// TIA Portal V19 export
// export: Created 2026-10-15T09:44:25.0424598Z, ExportSetting WithDefaults, DisplayName Totally Integrated Automation Portal, DisplayVersion V19, DisplayName TIA Portal Openness, DisplayVersion V19, DisplayName TIA Portal Version Control Interface, DisplayVersion V19, DisplayName STEP 7 Professional, DisplayVersion V19, DisplayName STEP 7 Safety, DisplayVersion V19, DisplayName WinCC Basic/Comfort/Advanced, DisplayVersion V19, DisplayName WinCC Unified, DisplayVersion V19
FUNCTION "ROLL_PB52" : Void   // FC35, SCL
{ S7_Optimized_Access := 'TRUE' }
VERSION : 0.1
// stored: AutoNumber true, IsIECCheckEnabled false, SetENOAutomatically false, UDAEnableTagReadback false
   VAR_TEMP
      r : Bool;
      a1 : Word;
      a2 : Word;
      activeDataBlock : Int;
      comparisonResults : Array[0..0] of Bool;
   END_VAR
BEGIN

   #r := FALSE;
   #a1 := W#16#0000;
   #a2 := W#16#0000;
   #activeDataBlock := 0;
   // PB52, STEP 5 network 1
   #activeDataBlock := 15;
   // PB52, STEP 5 network 2
   #a2 := #a1;
   #a1 := "ROLL_GetDW"(DbNumber := #activeDataBlock, Index := 17);
   #r := ((NOT "ROLL_IO".Input[5, 5]) AND (NOT "ROLL_State".M[6, 3]) AND "ROLL_IO".Input[3, 1] AND "ROLL_State".M[4, 1] AND "ROLL_State".M[40, 5]);
   "ROLL_TimerOp"(Number := 17,
                  Operation := 0,
                  Signal := #r,
                  Preset := #a1);
   // PB52, STEP 5 network 3
   #a2 := #a1;
   #a1 := "ROLL_GetDW"(DbNumber := #activeDataBlock, Index := 31);
   #r := ((NOT "ROLL_IO".Input[5, 3]) AND (NOT "ROLL_State".M[6, 1]) AND "ROLL_IO".Input[3, 1] AND "ROLL_State".M[4, 1]);
   "ROLL_TimerOp"(Number := 31,
                  Operation := 0,
                  Signal := #r,
                  Preset := #a1);
   // PB52, STEP 5 network 4
   #a2 := #a1;
   #a1 := "ROLL_GetDW"(DbNumber := #activeDataBlock, Index := 32);
   #r := ((NOT "ROLL_IO".Input[6, 0]) AND (NOT "ROLL_State".M[6, 4]) AND "ROLL_IO".Input[3, 1] AND "ROLL_State".M[4, 1]);
   "ROLL_TimerOp"(Number := 32,
                  Operation := 0,
                  Signal := #r,
                  Preset := #a1);
   // PB52, STEP 5 network 5
   #a2 := #a1;
   #a1 := "ROLL_GetDW"(DbNumber := #activeDataBlock, Index := 33);
   #r := ((NOT "ROLL_IO".Input[6, 2]) AND (NOT "ROLL_State".M[6, 5]) AND "ROLL_IO".Input[3, 1] AND "ROLL_State".M[4, 1]);
   "ROLL_TimerOp"(Number := 33,
                  Operation := 0,
                  Signal := #r,
                  Preset := #a1);
   // PB52, STEP 5 network 6
   #a2 := #a1;
   #a1 := W#16#3030;
   #r := ((NOT "ROLL_State".M[0, 4]) AND (NOT "ROLL_State".M[6, 7]) AND "ROLL_IO".Input[3, 1] AND "ROLL_State".M[4, 1]);
   "ROLL_TimerOp"(Number := 35,
                  Operation := 0,
                  Signal := #r,
                  Preset := #a1);
   // PB52, STEP 5 network 7
   #a2 := #a1;
   #a1 := W#16#3030;
   #r := ((NOT "ROLL_State".M[0, 4]) AND (NOT "ROLL_State".M[7, 0]) AND "ROLL_IO".Input[3, 1] AND "ROLL_State".M[4, 1]);
   "ROLL_TimerOp"(Number := 36,
                  Operation := 0,
                  Signal := #r,
                  Preset := #a1);
   // PB52, STEP 5 network 8
   #a2 := #a1;
   #a1 := W#16#3030;
   #r := ((NOT "ROLL_State".M[0, 4]) AND (NOT "ROLL_State".M[7, 1]) AND "ROLL_IO".Input[3, 1] AND "ROLL_State".M[4, 1]);
   "ROLL_TimerOp"(Number := 37,
                  Operation := 0,
                  Signal := #r,
                  Preset := #a1);
   // PB52, STEP 5 network 9
   #a2 := #a1;
   #a1 := W#16#3030;
   #r := ((NOT "ROLL_State".M[0, 4]) AND (NOT "ROLL_State".M[7, 2]) AND "ROLL_IO".Input[3, 1] AND "ROLL_State".M[4, 1]);
   "ROLL_TimerOp"(Number := 38,
                  Operation := 0,
                  Signal := #r,
                  Preset := #a1);
   // PB52, STEP 5 network 10
   #a2 := #a1;
   #a1 := W#16#1005;
   #r := "ROLL_IO".Input[123, 1];
   "ROLL_TimerOp"(Number := 45,
                  Operation := 0,
                  Signal := #r,
                  Preset := #a1);
   // PB52, STEP 5 network 11
   #a2 := #a1;
   #a1 := "ROLL_GetDW"(DbNumber := #activeDataBlock, Index := 58);
   #r := ("ROLL_IO".Input[3, 1] AND "ROLL_State".M[3, 6]);
   "ROLL_TimerOp"(Number := 58,
                  Operation := 1,
                  Signal := #r,
                  Preset := #a1);
   #a2 := #a1;
   #a1 := "ROLL_GetDW"(DbNumber := #activeDataBlock, Index := 59);
   #r := ("ROLL_State".M[3, 6] AND "ROLL_State".S5Timers[58].Q);
   "ROLL_TimerOp"(Number := 59,
                  Operation := 1,
                  Signal := #r,
                  Preset := #a1);
   // PB52, STEP 5 network 12
   #a2 := #a1;
   #a1 := "ROLL_GetDW"(DbNumber := #activeDataBlock, Index := 63);
   #r := (NOT "ROLL_State".S5Timers[62].Q);
   "ROLL_TimerOp"(Number := 63,
                  Operation := 0,
                  Signal := #r,
                  Preset := #a1);
   #a2 := #a1;
   #a1 := "ROLL_GetDW"(DbNumber := #activeDataBlock, Index := 62);
   #r := "ROLL_State".S5Timers[63].Q;
   "ROLL_TimerOp"(Number := 62,
                  Operation := 1,
                  Signal := #r,
                  Preset := #a1);
   #r := ((NOT "ROLL_State".M[103, 0]) AND (NOT "ROLL_State".M[103, 3]) AND (NOT "ROLL_State".M[103, 4]) AND (NOT "ROLL_State".S5Timers[119].Q));
   "ROLL_TimerOp"(Number := 62,
                  Operation := 2,
                  Signal := #r,
                  Preset := #a1);
   // PB52, STEP 5 network 13
   #a2 := #a1;
   #a1 := W#16#2010;
   #r := "ROLL_IO".Input[5, 3];
   "ROLL_TimerOp"(Number := 70,
                  Operation := 1,
                  Signal := #r,
                  Preset := #a1);
   // PB52, STEP 5 network 14
   #a2 := #a1;
   #a1 := W#16#2010;
   #r := "ROLL_IO".Input[6, 2];
   "ROLL_TimerOp"(Number := 72,
                  Operation := 1,
                  Signal := #r,
                  Preset := #a1);
   // PB52, STEP 5 network 15
   #a2 := #a1;
   #a1 := "ROLL_GetDW"(DbNumber := #activeDataBlock, Index := 85);
   #r := "ROLL_State".M[41, 0];
   "ROLL_TimerOp"(Number := 85,
                  Operation := 1,
                  Signal := #r,
                  Preset := #a1);
   // PB52, STEP 5 network 16
   RETURN;
END_FUNCTION
